(* IEC 61131-3 sources: kns-pump-station/tests/POUs/Station/FB_LevelControlPid_Test, 22 files *)

(* ---- AssistNotOffAboveAssistStartLevel.method.decl.st ---- *)
// 04 §7.2: при уровне не ниже 2,40 м подпорный не отключается даже при малом выходе ПИД — на всём интервале:
// без условия по уровню подпорный отключался бы через tAssistOff и снова включался по уровню через tLvlConfirm
// («качели»), а проверка только в конце интервала этого не видит
METHOD PRIVATE AssistNotOffAboveAssistStartLevel
VAR
    fbDut    : FB_LevelControlPid;          // ФБ под тестом
    fbTime   : PL.FB_FakeTime;              // подменное время, старт 1 ч
    stCfg    : ST_StationCfg;               // уставки по умолчанию (04 §18.2)
    afbPump  : ARRAY[1..3] OF FB_FakeMotorVfd;  // подменные насосы
    uiStep   : UINT;                        // шаг 100 мс
    xDropped : BOOL;                        // требуемое число хоть раз было не 2
END_VAR

(* ---- AssistNotOffAboveAssistStartLevel.method.impl.st ---- *)
coUnit.TEST('LevelPid_AssistNotOffAboveAssistStartLevel_A7');

fbDut.aitfPump[1] := afbPump[1];
fbDut.aitfPump[2] := afbPump[2];
fbDut.aitfPump[3] := afbPump[3];
fbDut.axCommOk[1] := TRUE;
fbDut.axCommOk[2] := TRUE;
fbDut.axCommOk[3] := TRUE;
fbDut.ePidMode := PL.E_DeviceMode.Auto;

afbPump[1].xRunning := TRUE;
afbPump[1].xSpeedAuto := TRUE;
afbPump[1].rSpeedRef := 60.0;
fbDut.uiLead := 1;
fbDut(xEnable := TRUE, rLevel_m := 2.5, xLevelValid := TRUE, rPidOut_pct := 50.0, xInit := TRUE,
      uiInitPumps := 2, itfTime := fbTime, stCfg := stCfg);

xDropped := FALSE;
FOR uiStep := 1 TO 1200 DO
    Run(fbDut := fbDut, fbTime := fbTime, stCfg := stCfg, rLevel_m := 2.5, rPidOut_pct := 50.0, uiSteps := 1);
    xDropped := xDropped OR fbDut.uiRequired <> 2;
END_FOR
AssertFalse(Condition := xDropped, Message := 'two pumps kept at 2.5 m for 120 s');

coUnit.TEST_FINISHED();

(* ---- AssistOffOutputLowForTAssistOff.method.decl.st ---- *)
// 04 §7.2, PMI-05: выход ПИД 75 % (граница включительно) дольше tAssistOff = 60 с при уровне ниже 2,40 м — один
// насос
METHOD PRIVATE AssistOffOutputLowForTAssistOff
VAR
    fbDut   : FB_LevelControlPid;           // ФБ под тестом
    fbTime  : PL.FB_FakeTime;               // подменное время, старт 1 ч
    stCfg   : ST_StationCfg;                // уставки по умолчанию (04 §18.2)
    afbPump : ARRAY[1..3] OF FB_FakeMotorVfd;   // подменные насосы
END_VAR

(* ---- AssistOnLevelAboveAssistStart.method.decl.st ---- *)
// 04 §7.2: уровень не ниже rLvlStartAssist_m = 2,40 м дольше tLvlConfirm — второй насос и при малом выходе ПИД
METHOD PRIVATE AssistOnLevelAboveAssistStart
VAR
    fbDut   : FB_LevelControlPid;           // ФБ под тестом
    fbTime  : PL.FB_FakeTime;               // подменное время, старт 1 ч
    stCfg   : ST_StationCfg;                // уставки по умолчанию (04 §18.2)
    afbPump : ARRAY[1..3] OF FB_FakeMotorVfd;   // подменные насосы
END_VAR

(* ---- AssistOnOutputHighForTAssistOn.method.decl.st ---- *)
// 04 §7.2, PMI-05: выход ПИД 98 % (граница включительно) дольше tAssistOn = 30 с — второй насос, не раньше
METHOD PRIVATE AssistOnOutputHighForTAssistOn
VAR
    fbDut   : FB_LevelControlPid;           // ФБ под тестом
    fbTime  : PL.FB_FakeTime;               // подменное время, старт 1 ч
    stCfg   : ST_StationCfg;                // уставки по умолчанию (04 §18.2)
    afbPump : ARRAY[1..3] OF FB_FakeMotorVfd;   // подменные насосы
END_VAR

(* ---- CommAbsentDuringPowerRestoreNoRecoverDelay.method.decl.st ---- *)
// 04 §7.4, §12, §13, VFD-12 plc-process-lib: напряжение восстановлено, насосы доступны, а ПЧ ещё загружаются
// (связи нет) — это не потеря связи: выдержка возврата STN_PID_RECOVER не перезапускается, ПИД готов, как только
// связь появилась. Вне окна восстановления питания прежнее правило: связь пропала у всех — возврат через 30 с
METHOD PRIVATE CommAbsentDuringPowerRestoreNoRecoverDelay
VAR
    fbDut   : FB_LevelControlPid;           // ФБ под тестом
    fbTime  : PL.FB_FakeTime;               // подменное время, старт 1 ч
    stCfg   : ST_StationCfg;                // уставки по умолчанию (04 §18.2)
    afbPump : ARRAY[1..3] OF FB_FakeMotorVfd;   // подменные насосы: доступны, Auto, стоят
    uiStep  : UINT;                         // шаг 100 мс
    uiIdx   : UINT;                         // насос
END_VAR

(* ---- CommAbsentDuringPowerRestoreNoRecoverDelay.method.impl.st ---- *)
coUnit.TEST('LevelPid_CommAbsentDuringPowerRestoreNoRecoverDelay_A7_A12_A13');

fbDut.aitfPump[1] := afbPump[1];
fbDut.aitfPump[2] := afbPump[2];
fbDut.aitfPump[3] := afbPump[3];
fbDut.axCommOk[1] := TRUE;
fbDut.axCommOk[2] := TRUE;
fbDut.axCommOk[3] := TRUE;
fbDut.ePidMode := PL.E_DeviceMode.Auto;
fbDut(xEnable := FALSE, rLevel_m := 1.2, xLevelValid := TRUE, itfTime := fbTime, stCfg := stCfg);
AssertTrue(Condition := fbDut.xPidReady, Message := 'stopped pumps with comm: ready');

// нет напряжения: насосы недоступны, ПЧ без питания — связи нет
fbDut.xPowerRestore := TRUE;
FOR uiIdx := 1 TO 3 DO
    afbPump[uiIdx].xAvailable := FALSE;
    fbDut.axCommOk[uiIdx] := FALSE;
END_FOR
FOR uiStep := 1 TO 100 DO
    fbTime.Advance(tStep := T#100MS);
    fbDut(xEnable := FALSE, itfTime := fbTime, stCfg := stCfg);
END_FOR
AssertFalse(Condition := fbDut.xPidReady, Message := 'power lost: not ready');
// напряжение восстановлено: насосы доступны, ПЧ 2 с загружаются
FOR uiIdx := 1 TO 3 DO
    afbPump[uiIdx].xAvailable := TRUE;
END_FOR
FOR uiStep := 1 TO 20 DO
    fbTime.Advance(tStep := T#100MS);
    fbDut(xEnable := FALSE, itfTime := fbTime, stCfg := stCfg);
END_FOR
AssertFalse(Condition := fbDut.xPidReady, Message := 'drives booting: not ready');
fbDut.axCommOk[1] := TRUE;
fbTime.Advance(tStep := T#100MS);
fbDut(xEnable := FALSE, itfTime := fbTime, stCfg := stCfg);
AssertTrue(Condition := fbDut.xPidReady, Message := 'drive booted: ready at once, no recover delay');

// после восстановления питания: связь пропала у всех — снова через STN_PID_RECOVER
fbDut.xPowerRestore := FALSE;
fbDut.axCommOk[1] := FALSE;
fbTime.Advance(tStep := T#100MS);
fbDut(xEnable := FALSE, itfTime := fbTime, stCfg := stCfg);
AssertFalse(Condition := fbDut.xPidReady, Message := 'comm lost outside power restore: not ready');
fbDut.axCommOk[1] := TRUE;
FOR uiStep := 1 TO 300 DO
    fbTime.Advance(tStep := T#100MS);
    fbDut(xEnable := FALSE, itfTime := fbTime, stCfg := stCfg);
END_FOR
AssertFalse(Condition := fbDut.xPidReady, Message := 'not ready 29.9 s after comm recovery');
fbTime.Advance(tStep := T#100MS);
fbDut(xEnable := FALSE, itfTime := fbTime, stCfg := stCfg);
AssertTrue(Condition := fbDut.xPidReady, Message := 'ready 30 s after comm recovery');

coUnit.TEST_FINISHED();

(* ---- HoldOutputWhenLeadDropsOut.method.decl.st ---- *)
// 04 §7.3, §9: ведущий прошлого цикла выбыл (авария ПЧ, блокировка станции) при выбранном ПИД — выход ПИД
// держится (слежение за собственным выходом), а не за заданием 0 выбывшего ПЧ; ПИД не выбран или ведущий доступен
// (пуск) — слежение за заданием ведущего, как раньше
METHOD PRIVATE HoldOutputWhenLeadDropsOut
VAR
    fbDut   : FB_LevelControlPid;           // ФБ под тестом
    fbTime  : PL.FB_FakeTime;               // подменное время, старт 1 ч
    stCfg   : ST_StationCfg;                // уставки по умолчанию (04 §18.2)
    afbPump : ARRAY[1..3] OF FB_FakeMotorVfd;   // подменные насосы
END_VAR

(* ---- InitFromRunningPumps.method.decl.st ---- *)
// 04 §3.2, PMI-07: вход без рывка — число насосов по работающим, не больше MIN(2, uiDutyMax)
METHOD PRIVATE InitFromRunningPumps
VAR
    fbDut   : FB_LevelControlPid;           // ФБ под тестом
    fbTime  : PL.FB_FakeTime;               // подменное время, старт 1 ч
    stCfg   : ST_StationCfg;                // уставки по умолчанию (04 §18.2)
    afbPump : ARRAY[1..3] OF FB_FakeMotorVfd;   // подменные насосы
    fbDut2  : FB_LevelControlPid;          // второй экземпляр: uiDutyMax = 1
    stCfg1  : ST_StationCfg;               // уставки с uiDutyMax = 1
END_VAR

(* ---- NanOutputNoStaging.method.decl.st ---- *)
// Неконечный выход ПИД — подключение и отключение подпорного по выходу не срабатывают (сравнения с NaN ложны)
METHOD PRIVATE NanOutputNoStaging
VAR
    fbDut   : FB_LevelControlPid;           // ФБ под тестом
    fbTime  : PL.FB_FakeTime;               // подменное время, старт 1 ч
    stCfg   : ST_StationCfg;                // уставки по умолчанию (04 §18.2)
    afbPump : ARRAY[1..3] OF FB_FakeMotorVfd;   // подменные насосы
    rNan    : REAL;                     // NaN
    uBits   : PL.U_RealBits;             // сборка NaN по битам
    fbDut2  : FB_LevelControlPid;          // второй экземпляр: два насоса
END_VAR

(* ---- NotReadyWhenPidManual.method.decl.st ---- *)
// 04 §7.4: ПИД не в Auto или уровень негоден — не готов
METHOD PRIVATE NotReadyWhenPidManual
VAR
    fbDut   : FB_LevelControlPid;           // ФБ под тестом
    fbTime  : PL.FB_FakeTime;               // подменное время, старт 1 ч
    stCfg   : ST_StationCfg;                // уставки по умолчанию (04 §18.2)
    afbPump : ARRAY[1..3] OF FB_FakeMotorVfd;   // подменные насосы
END_VAR

(* ---- NotReadyWithoutCommPump.method.decl.st ---- *)
// 04 §7.4, PMI-29: нет насоса со связью — ни среди работающих, ни среди доступных стоящих — ПИД не готов
METHOD PRIVATE NotReadyWithoutCommPump
VAR
    fbDut   : FB_LevelControlPid;           // ФБ под тестом
    fbTime  : PL.FB_FakeTime;               // подменное время, старт 1 ч
    stCfg   : ST_StationCfg;                // уставки по умолчанию (04 §18.2)
    afbPump : ARRAY[1..3] OF FB_FakeMotorVfd;   // подменные насосы
END_VAR

(* ---- OutputStagingOnlyWhenPidControls.method.decl.st ---- *)
// Условия по выходу ПИД действуют, только когда ПИД управляет: выход 100 % в слежении (ведущий не в
// SpeedAutoActive) подпорного не включает
METHOD PRIVATE OutputStagingOnlyWhenPidControls
VAR
    fbDut   : FB_LevelControlPid;           // ФБ под тестом
    fbTime  : PL.FB_FakeTime;               // подменное время, старт 1 ч
    stCfg   : ST_StationCfg;                // уставки по умолчанию (04 §18.2)
    afbPump : ARRAY[1..3] OF FB_FakeMotorVfd;   // подменные насосы
END_VAR

(* ---- ReadyAfterCommRecoverDelay.method.decl.st ---- *)
// 04 §12, PMI-28: связь пропала у всех — готовность снимается сразу; вернулась — готовность через STN_PID_RECOVER
// = 30 с, не раньше
METHOD PRIVATE ReadyAfterCommRecoverDelay
VAR
    fbDut   : FB_LevelControlPid;           // ФБ под тестом
    fbTime  : PL.FB_FakeTime;               // подменное время, старт 1 ч
    stCfg   : ST_StationCfg;                // уставки по умолчанию (04 §18.2)
    afbPump : ARRAY[1..3] OF FB_FakeMotorVfd;   // подменные насосы
    uiStep  : UINT;                     // шаг 100 мс
END_VAR

(* ---- ReadyAfterCommRecoverDelay.method.impl.st ---- *)
coUnit.TEST('LevelPid_ReadyAfterCommRecoverDelay_A7_A12_PMI28');

fbDut.aitfPump[1] := afbPump[1];
fbDut.aitfPump[2] := afbPump[2];
fbDut.aitfPump[3] := afbPump[3];
fbDut.axCommOk[1] := TRUE;
fbDut.axCommOk[2] := TRUE;
fbDut.axCommOk[3] := TRUE;
fbDut.ePidMode := PL.E_DeviceMode.Auto;

afbPump[1].xRunning := TRUE;
afbPump[1].xSpeedAuto := TRUE;
afbPump[1].rSpeedRef := 60.0;
fbDut.uiLead := 1;

fbDut(xEnable := TRUE, rLevel_m := 1.5, xLevelValid := TRUE, itfTime := fbTime, stCfg := stCfg);
AssertTrue(Condition := fbDut.xPidReady, Message := 'running pump with comm: ready');
fbDut.axCommOk[1] := FALSE;
fbDut.axCommOk[2] := FALSE;
fbDut.axCommOk[3] := FALSE;
fbTime.Advance(tStep := T#100MS);
fbDut(xEnable := TRUE, itfTime := fbTime, stCfg := stCfg);
AssertFalse(Condition := fbDut.xPidReady, Message := 'comm lost: not ready at once');
fbDut.axCommOk[1] := TRUE;
FOR uiStep := 1 TO 300 DO
    fbTime.Advance(tStep := T#100MS);
    fbDut(xEnable := TRUE, itfTime := fbTime, stCfg := stCfg);
END_FOR
AssertFalse(Condition := fbDut.xPidReady, Message := 'not ready 29.9 s after comm recovery');
fbTime.Advance(tStep := T#100MS);
fbDut(xEnable := TRUE, itfTime := fbTime, stCfg := stCfg);
AssertTrue(Condition := fbDut.xPidReady, Message := 'ready 30 s after comm recovery');

coUnit.TEST_FINISHED();

(* ---- Run.method.decl.st ---- *)
// Помощник: uiSteps шагов по 100 мс с одним уровнем и выходом ПИД (ПИД выбран, уровень достоверен)
METHOD PRIVATE Run
VAR_IN_OUT
    fbDut  : FB_LevelControlPid;        // ФБ под тестом
    fbTime : PL.FB_FakeTime;            // подменное время
    stCfg  : ST_StationCfg;             // уставки
END_VAR
VAR_INPUT
    rLevel_m    : REAL;                 // уровень
    rPidOut_pct : REAL;                 // выход ПИД
    uiSteps     : UINT;                 // шагов по 100 мс
END_VAR
VAR
    uiStep : UINT;                      // номер шага
END_VAR

(* ---- Run.method.impl.st ---- *)
FOR uiStep := 1 TO uiSteps DO
    fbTime.Advance(tStep := T#100MS);
    fbDut(xEnable := TRUE, rLevel_m := rLevel_m, xLevelValid := TRUE, rPidOut_pct := rPidOut_pct, xInit := FALSE,
          itfTime := fbTime, stCfg := stCfg);
END_FOR

(* ---- StartsLeadAtStartLevel.method.decl.st ---- *)
// 04 §7.2, PMI-04: насосы стоят, уровень 1,60 м — пуск ведущего через tLvlConfirm = 5 с
METHOD PRIVATE StartsLeadAtStartLevel
VAR
    fbDut   : FB_LevelControlPid;           // ФБ под тестом
    fbTime  : PL.FB_FakeTime;               // подменное время, старт 1 ч
    stCfg   : ST_StationCfg;                // уставки по умолчанию (04 §18.2)
    afbPump : ARRAY[1..3] OF FB_FakeMotorVfd;   // подменные насосы
END_VAR

(* ---- StopAllAtStopLevel.method.decl.st ---- *)
// 04 §7.2, PMI-06: уровень 1,00 м дольше tLvlConfirm — все насосы стоп, в том числе из двух
METHOD PRIVATE StopAllAtStopLevel
VAR
    fbDut   : FB_LevelControlPid;           // ФБ под тестом
    fbTime  : PL.FB_FakeTime;               // подменное время, старт 1 ч
    stCfg   : ST_StationCfg;                // уставки по умолчанию (04 §18.2)
    afbPump : ARRAY[1..3] OF FB_FakeMotorVfd;   // подменные насосы
END_VAR

(* ---- TimeBackwardsRestartsConfirm.method.decl.st ---- *)
// Время назад (сбой источника) — выдержка подтверждения пуска ведущего начинается заново, ложного пуска нет
METHOD PRIVATE TimeBackwardsRestartsConfirm
VAR
    fbDut   : FB_LevelControlPid;           // ФБ под тестом
    fbTime  : PL.FB_FakeTime;               // подменное время, старт 1 ч
    stCfg   : ST_StationCfg;                // уставки по умолчанию (04 §18.2)
    afbPump : ARRAY[1..3] OF FB_FakeMotorVfd;   // подменные насосы
END_VAR

(* ---- TrackWhenLeadCommLost.method.decl.st ---- *)
// 04 §12, PMI-28: у ведущего нет связи с ПЧ — ПИД в слежении (интегратор не копится против замершей частоты)
METHOD PRIVATE TrackWhenLeadCommLost
VAR
    fbDut   : FB_LevelControlPid;           // ФБ под тестом
    fbTime  : PL.FB_FakeTime;               // подменное время, старт 1 ч
    stCfg   : ST_StationCfg;                // уставки по умолчанию (04 §18.2)
    afbPump : ARRAY[1..3] OF FB_FakeMotorVfd;   // подменные насосы
END_VAR

(* ---- TrackWhenLeadNotSpeedAuto.method.decl.st ---- *)
// 04 §7.3, PMI-04: ведущий работает, но не в SpeedAutoActive — ПИД в слежении за его заданием; ведущего нет —
// слежение за 0
METHOD PRIVATE TrackWhenLeadNotSpeedAuto
VAR
    fbDut   : FB_LevelControlPid;           // ФБ под тестом
    fbTime  : PL.FB_FakeTime;               // подменное время, старт 1 ч
    stCfg   : ST_StationCfg;                // уставки по умолчанию (04 §18.2)
    afbPump : ARRAY[1..3] OF FB_FakeMotorVfd;   // подменные насосы
END_VAR
